PROGRAM main
  VAR
    S1 AT %IX0.0  : BOOL; (* marcha / lote nuevo, NA *)
    S0 AT %IX0.1  : BOOL; (* parada, NC: TRUE sin pulsar *)
    B1 AT %IX0.2  : BOOL; (* sensor de piezas *)
    KM1 AT %QX0.0 : BOOL; (* motor de la cinta *)
    H1 AT %QX0.1  : BOOL; (* lote completo *)
    F_PIEZA       : R_TRIG;
    PIEZA         : BOOL; (* flanco de B1 *)
    PIEZAS        : INT; (* piezas del lote *)
    COMPLETO      : BOOL; (* lote completo *)
    F_LOTE        : R_TRIG;
    LOTE_NUEVO    : BOOL; (* flanco de COMPLETO *)
    LOTES         : INT; (* lotes completos en el turno *)
    TURNO         : BOOL; (* turno completo *)
  END_VAR
  VAR  (* added by the conversion: wires and edge detectors of the diagram *)
    _AND5_OUT : BOOL;
    _ADD9_OUT : INT;
    _SEL4_OUT : INT;
    _AND14_OUT : BOOL;
    _SEL13_OUT : INT;
    _GE20_OUT : BOOL;
    _OR25_OUT : BOOL;
    _NOT29_OUT : BOOL;
    _AND24_OUT : BOOL;
  END_VAR

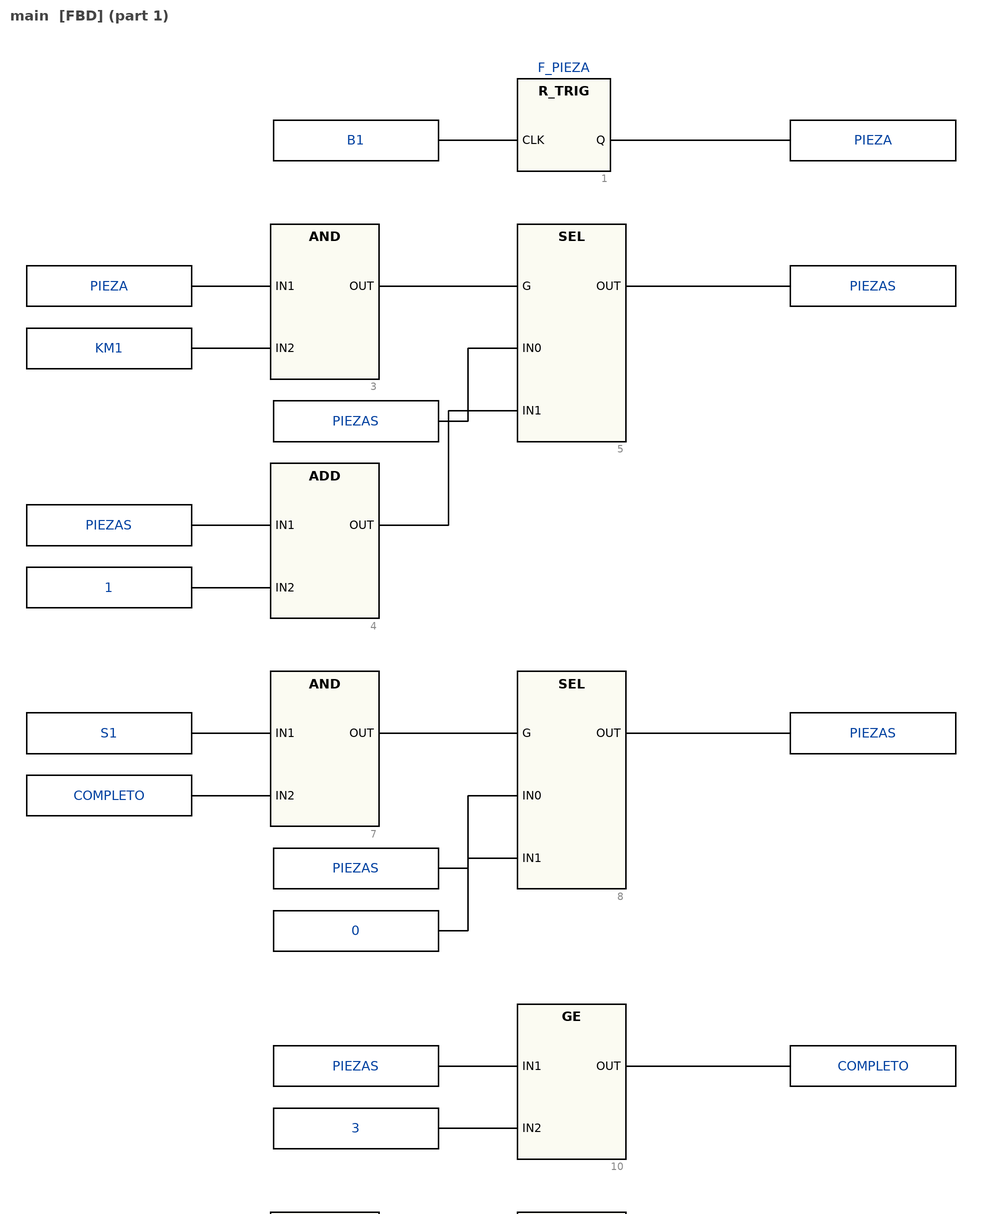
(* FBD diagram, written out as Structured Text *)
F_PIEZA(CLK := B1);
PIEZA := F_PIEZA.Q;
_AND5_OUT := PIEZA AND KM1;
_ADD9_OUT := PIEZAS + 1;
_SEL4_OUT := SEL(_AND5_OUT, PIEZAS, _ADD9_OUT);
PIEZAS := _SEL4_OUT;
_AND14_OUT := S1 AND COMPLETO;
_SEL13_OUT := SEL(_AND14_OUT, PIEZAS, 0);
PIEZAS := _SEL13_OUT;
_GE20_OUT := PIEZAS >= 3;
COMPLETO := _GE20_OUT;
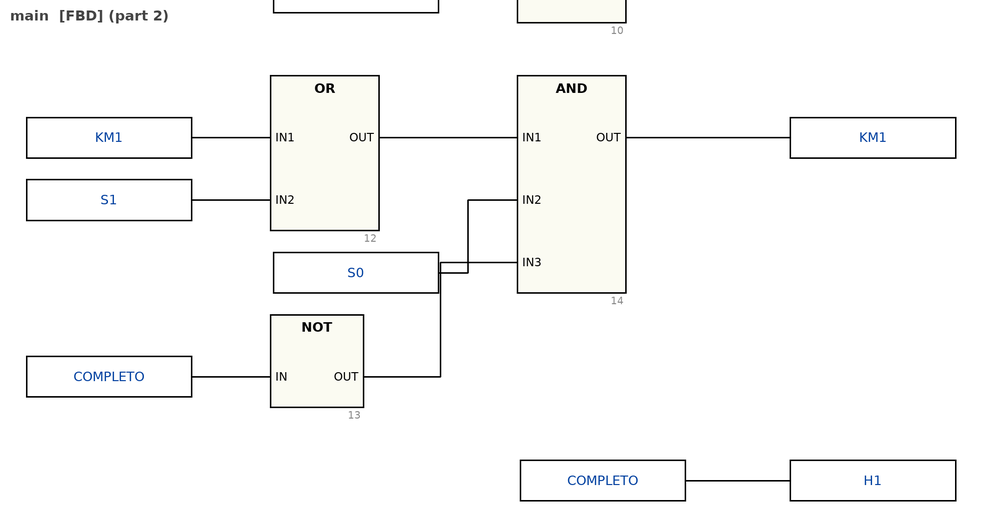
_OR25_OUT := KM1 OR S1;
_NOT29_OUT := NOT COMPLETO;
_AND24_OUT := _OR25_OUT AND S0 AND _NOT29_OUT;
KM1 := _AND24_OUT;
H1 := COMPLETO;
END_PROGRAM
